Fanuc KAREL source: kb00157.KL

-- PROVISIONAL review KL for V1013-1; original PC SHA256 a7525ef2c5c5c07dfc04269614148110a2384af060723fad653a88469bfbbfba
-- Incomplete behavior may be omitted. Consult companion uncertainty JSON. Do not deploy.
PROGRAM KB00157
%NOLOCKGROUP
BEGIN
  -- UNRESOLVED_PC offsets 5-12; opcodes 9D,23
  -- UNRESOLVED_PC offsets 17-33; opcodes 27,22,31,23
  -- UNRESOLVED_PC offsets 38-42; opcodes 7F
END KB00157
